FUNCTION_BLOCK FB_Jog_Joint
VAR_INPUT
	// Misc:
	lr_DeltaTime : LREAL;
	
	// Config parameters
	lr_SlowModeVelocitySetting : LREAL; // [deg/s]
	lr_FastModeVelovitySetting : LREAL; // [deg/s]
	i_Base_LowLimit : INT;
	i_Base_HighLimit : INT;
	i_Shoulder_LowLimit : INT;
	i_Shoulder_HighLimit : INT;
	i_Elbow_LowLimit : INT;
	i_Elbow_HighLimit : INT;
	
	
	
	// Control inputs
	b_Enable_Servos : BOOL;
	SW_Fast_Mode : BOOL; // True = fast mode, False = slow mode
	PB_Base_Pos : BOOL;
	PB_Base_Neg : BOOL;
	PB_Shoulder_Pos : BOOL;
	PB_Shoulder_Neg : BOOL;
	PB_Elbow_Pos : BOOL;
	PB_Elbow_Neg : BOOL;


END_VAR
VAR_OUTPUT
	i_Set_Base : INT;
	i_Set_Shoulder : INT;
	i_Set_Elbow : INT;
END_VAR
VAR
	lr_CurrentSpeedSetting : LREAL; // [deg/s]
	lr_Set_Base : LREAL;
	lr_Set_Shoulder : LREAL;
	lr_Set_Elbow : LREAL;
	
		// Structures:
	fb_Servo_Base : FB_Servo;
	fb_Servo_Shoulder : FB_Servo;
	fb_Servo_Elbow : FB_Servo;
END_VAR

fb_Servo_Base(
	b_EnableServo:= b_Enable_Servos, 
	b_CW:= PB_Base_Neg, 
	b_CCW:= PB_Base_Pos, 
	lr_deltaTime:= lr_DeltaTime, 
	lr_DegLowLim:= i_Base_LowLimit, 
	lr_DegHighLim:= i_Base_HighLimit, 
	lr_SlowModeVelocitySetting:= lr_SlowModeVelocitySetting, 
	lr_FastModeVelovitySetting:= lr_FastModeVelovitySetting, 
	SW_Fast_Mode:= SW_Fast_Mode, 
	i_Set_Angle=> i_Set_Base);

fb_Servo_Elbow(
	b_EnableServo:= b_Enable_Servos, 
	b_CW:= PB_Shoulder_Pos, 
	b_CCW:= PB_Shoulder_Neg, 
	lr_deltaTime:= lr_DeltaTime, 
	lr_DegLowLim:= i_Shoulder_LowLimit, 
	lr_DegHighLim:= i_Shoulder_HighLimit, 
	lr_SlowModeVelocitySetting:= lr_SlowModeVelocitySetting, 
	lr_FastModeVelovitySetting:= lr_FastModeVelovitySetting, 
	SW_Fast_Mode:= SW_Fast_Mode, 
	i_Set_Angle=> i_Set_Shoulder);

fb_Servo_Shoulder(
	b_EnableServo:= b_Enable_Servos, 
	b_CW:= PB_Elbow_Pos, 
	b_CCW:= PB_Elbow_Neg, 
	lr_deltaTime:= lr_DeltaTime, 
	lr_DegLowLim:= i_Elbow_LowLimit, 
	lr_DegHighLim:= i_Elbow_HighLimit, 
	lr_SlowModeVelocitySetting:= lr_SlowModeVelocitySetting, 
	lr_FastModeVelovitySetting:= lr_FastModeVelovitySetting, 
	SW_Fast_Mode:= SW_Fast_Mode, 
	i_Set_Angle=> i_Set_Elbow);

END_FUNCTION_BLOCK

(* stored: Version 1.1.0.1, ProductVersion 3.1.4024.13
   POU FB_Jog_Joint: Id {52a44315-b2e5-4aeb-9b6c-90503662b0b6}, SpecialFunc None *)
